SUBAPPLICATION Servo_AI3_Calibrate_2P_OPC (* Servo an Output_Q2 folgt dem 2-Punkt-kalibrierten Slider AI3 (0-180 Grad), Kalibrierung CO/CS + Referenzwerte per OPC-UA-Dashboard *)
  (* Standard: 61499-2; Description: Copyright (c) 2026 Meisterschulen am Ostbahnhof This program and the accompanying materials are made available under the terms of the Eclipse Public License 2.0 which is available at https://www.eclipse.org/legal/epl-2.0/ SPDX-License-Identifier: EPL-2.0 *)
  (* Version 1.0, 2026-11-06, Franz Höpfinger, Meisterschulen am Ostbahnhof, Kopie von Meins::Servo_AI4_Calibrate_OPC fuer den Slider AI3 (haelt seine Position, keine Mittelstellung): 2-Punkt-Kalibrierung MyLib::sys::logiBUS_AI_Calibrate_2P_OPC statt 3P. Kalibrierter Wert = Winkel in Grad, Referenzwerte 0/180. *)
  PACKAGE Meins::Servo_AI3_Calibrate_2P_OPC;
  IMPORT Meins::Servo_AI3_Calibrate_2P_OPC::SubStrings::SAI3_RAW_WRITE;
  IMPORT Meins::Servo_AI3_Calibrate_2P_OPC::SubStrings::SAI3_CAL_WRITE;
  IMPORT Meins::Servo_AI3_Calibrate_2P_OPC::SubStrings::SAI3_CO_METHOD;
  IMPORT Meins::Servo_AI3_Calibrate_2P_OPC::SubStrings::SAI3_CS_METHOD;
  IMPORT Meins::Servo_AI3_Calibrate_2P_OPC::SubStrings::SAI3_ZERO_READ;
  IMPORT Meins::Servo_AI3_Calibrate_2P_OPC::SubStrings::SAI3_ZERO_WRITE;
  IMPORT Meins::Servo_AI3_Calibrate_2P_OPC::SubStrings::SAI3_SPAN_READ;
  IMPORT Meins::Servo_AI3_Calibrate_2P_OPC::SubStrings::SAI3_SPAN_WRITE;
  IMPORT Meins::Servo_AI3_Calibrate_2P_OPC::SubStrings::SAI3_ZERO_RAW_WRITE;
  IMPORT Meins::Servo_AI3_Calibrate_2P_OPC::SubStrings::SAI3_SPAN_RAW_WRITE;
  IMPORT Meins::Servo_AI3_Calibrate_2P_OPC::SubStrings::SAI3_ANGLE;
  IMPORT logiBUS::io::AI::logiBUS_AI::AnalogInput_I3;
  IMPORT logiBUS::io::DQ::logiBUS_DO::Output_Q2;
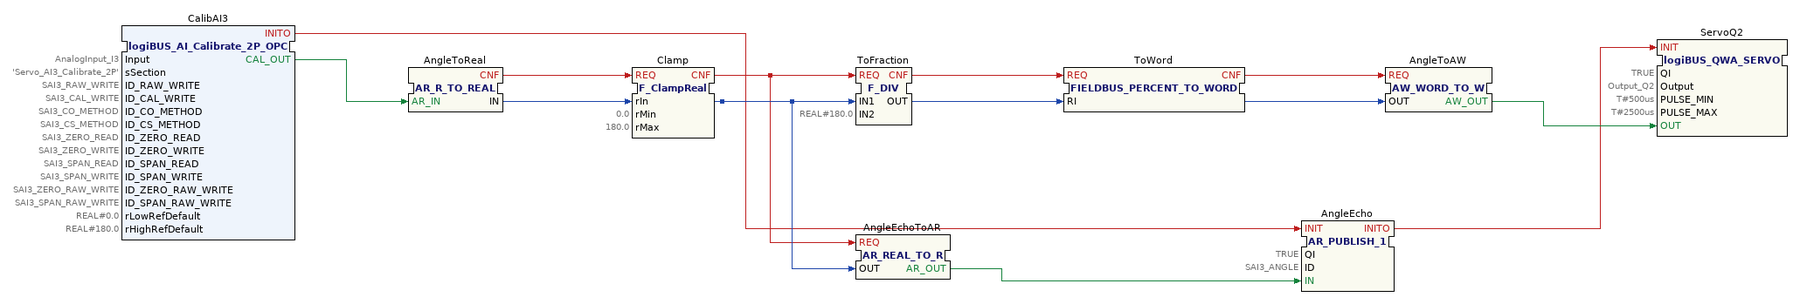
  (* ServoQ2: PULSE_MIN = T#500us, PULSE_MAX = T#2500us, FREQ 50 Hz (Mitte 1,5 ms). Passt fuer: 5 Stueck 9G Servo Motor, Mikro-Servomotoren mit Kabel, 180 Grad (Amazon B0H3BC3PSS). Herstellerangabe: 20 ms Zyklus, 0,5..2,5 ms Impulsbreite fuer 0..180 Grad, 3..7,2 V. Damit faehrt der Servo exakt 90 Grad in jede Richtung (getestet 2026-11-06). Standardwerte 1000..2000 us ergeben bei diesem Servo nur ca. 35 Grad. *)
  FBS
    AngleToReal : adapter::conversion::unidirectional::AR_R_TO_REAL;
    Clamp : logiBUS::signalprocessing::clamp::F_ClampReal(rMin := 0.0, rMax := 180.0);
    ToFraction : iec61131::arithmetic::F_DIV(IN2 := REAL#180.0);
    ToWord : eclipse4diac::signalprocessing::FIELDBUS_PERCENT_TO_WORD;
    AngleToAW : adapter::conversion::unidirectional::AW_WORD_TO_W;
    ServoQ2 : logiBUS::io::DO_SERVO::logiBUS_QWA_SERVO(QI := TRUE, Output := Output_Q2, PULSE_MIN := T#500us, PULSE_MAX := T#2500us);
    AngleEchoToAR : adapter::conversion::unidirectional::AR_REAL_TO_R;
    AngleEcho : adapter::net::AR_PUBLISH_1(QI := TRUE, ID := SAI3_ANGLE);
  END_FBS
  SUBAPPS
    CalibAI3 : MyLib::sys::logiBUS_AI_Calibrate_2P_OPC(Input := AnalogInput_I3, sSection := 'Servo_AI3_Calibrate_2P', ID_RAW_WRITE := SAI3_RAW_WRITE, ID_CAL_WRITE := SAI3_CAL_WRITE, ID_CO_METHOD := SAI3_CO_METHOD, ID_CS_METHOD := SAI3_CS_METHOD, ID_ZERO_READ := SAI3_ZERO_READ, ID_ZERO_WRITE := SAI3_ZERO_WRITE, ID_SPAN_READ := SAI3_SPAN_READ, ID_SPAN_WRITE := SAI3_SPAN_WRITE, ID_ZERO_RAW_WRITE := SAI3_ZERO_RAW_WRITE, ID_SPAN_RAW_WRITE := SAI3_SPAN_RAW_WRITE, rLowRefDefault := REAL#0.0, rHighRefDefault := REAL#180.0);
  END_SUBAPPS
  EVENT_CONNECTIONS
    AngleToReal.CNF TO Clamp.REQ;
    Clamp.CNF TO ToFraction.REQ;
    Clamp.CNF TO AngleEchoToAR.REQ;
    ToFraction.CNF TO ToWord.REQ;
    ToWord.CNF TO AngleToAW.REQ;
    CalibAI3.INITO TO AngleEcho.INIT;
    AngleEcho.INITO TO ServoQ2.INIT;
  END_CONNECTIONS
  DATA_CONNECTIONS
    AngleToReal.IN TO Clamp.rIn;
    Clamp. TO ToFraction.IN1;
    ToFraction.OUT TO ToWord.RI;
    ToWord. TO AngleToAW.OUT;
    Clamp. TO AngleEchoToAR.OUT;
  END_CONNECTIONS
  ADAPTER_CONNECTIONS
    CalibAI3.CAL_OUT TO AngleToReal.AR_IN;
    AngleToAW.AW_OUT TO ServoQ2.OUT;
    AngleEchoToAR.AR_OUT TO AngleEcho.IN;
  END_CONNECTIONS
END_SUBAPPLICATION
